Fanuc KAREL source: KT00536.KL

PROGRAM KT00536
%NOLOCKGROUP
VAR
  P1: JOINTPOS
  P2: POSITION
  OUT: XYZWPREXT
BEGIN
  OUT = P1 : P2
END KT00536
